Staubli VAL3: _clickFuncReset.pgx

public program _clickFuncReset()
  local num l_nI
begin
  //“全部复位”按钮回调（无参数，供 AppStart.bindings.json 的 callbacks 调用）
  //9 个功能按钮选中态清零，背景色回默认灰
  for l_nI=0 to 8
    bFunc[l_nI]=false
    sFuncBg[l_nI]="#DCDCDC"
  endFor
end
